FUNCTION_BLOCK F (* Needs reading R3: exit guards after a shared algorithm that only sometimes assigns, so the value read may be the carried-over one *)
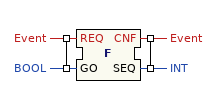
  EVENT_INPUT
    REQ WITH GO;
  END_EVENT
  EVENT_OUTPUT
    CNF WITH SEQ;
  END_EVENT
  VAR_INPUT
    GO : BOOL;
  END_VAR
  VAR_OUTPUT
    SEQ : INT;
  END_VAR
  VAR
    D : INT;
  END_VAR
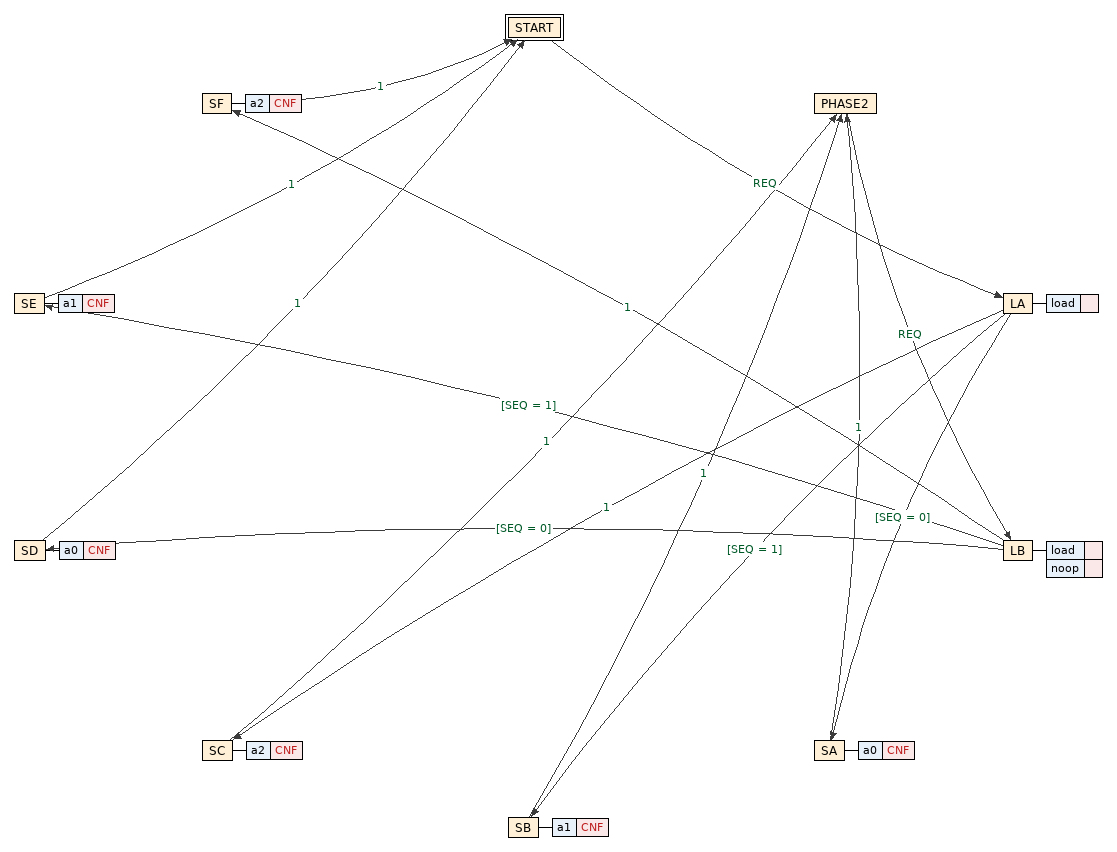
  EC_STATES
    START;
    PHASE2;
    LA : load;
    LB : load, noop;
    SA : a0 -> CNF;
    SB : a1 -> CNF;
    SC : a2 -> CNF;
    SD : a0 -> CNF;
    SE : a1 -> CNF;
    SF : a2 -> CNF;
  END_STATES
  EC_TRANSITIONS
    START TO LA := REQ;
    PHASE2 TO LB := REQ;
    LA TO SA := [SEQ = 0];
    LA TO SB := [SEQ = 1];
    LA TO SC := 1;
    LB TO SD := [SEQ = 0];
    LB TO SE := [SEQ = 1];
    LB TO SF := 1;
    SA TO PHASE2 := 1;
    SB TO PHASE2 := 1;
    SC TO PHASE2 := 1;
    SD TO START := 1;
    SE TO START := 1;
    SF TO START := 1;
  END_TRANSITIONS
  ALGORITHM load IN ST:
IF GO THEN
  SEQ := 2;
END_IF;
  END_ALGORITHM
  ALGORITHM a0 IN ST:
SEQ := 1;
  END_ALGORITHM
  ALGORITHM a1 IN ST:
SEQ := 2;
  END_ALGORITHM
  ALGORITHM a2 IN ST:
SEQ := 0;
  END_ALGORITHM
  ALGORITHM noop IN ST:
D := 0;
  END_ALGORITHM
END_FUNCTION_BLOCK
